INTERFACE PUBLIC Drive EXTENDS __System.IQueryInterface

END_INTERFACE

(* stored: Version 1.1.0.1
   Itf Drive: Id {bf1dd6ff-2760-40cd-9171-687ef61d1525} *)
